FUNCTION_BLOCK logiBUS_QWA_SERVO (* Composite FB for servo word output data *)
  (* Standard: 61499-2; Description: Copyright (c) 2026 HR Agrartechnik GmbH This program and the accompanying materials are made available under the terms of the Eclipse Public License 2.0 which is available at https://www.eclipse.org/legal/epl-2.0/ SPDX-License-Identifier: EPL-2.0 *)
  (* Version 1.1, 2026-11-06, Franz Höpfinger, HR Agrartechnik GmbH, Servo on MCPWM with FREQ, PULSE_MIN, PULSE_MAX (before: LEDC, fixed 250 Hz, 800..2180 us) *)
  (* Version 1.0, 2026-02-23, Franz Höpfinger, HR Agrartechnik GmbH *)
  PACKAGE logiBUS::io::DO_SERVO;
  IMPORT logiBUS::io::DQ::logiBUS_DO::Invalid;
  IMPORT logiBUS::io::DQ::logiBUS_DO_S;
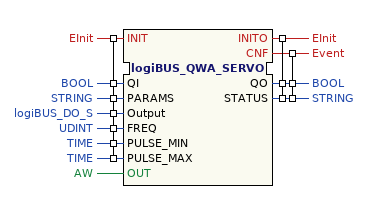
  EVENT_INPUT
    INIT : EInit WITH QI, PARAMS, Output, FREQ, PULSE_MIN, PULSE_MAX; (* Service Initialization *)
  END_EVENT
  EVENT_OUTPUT
    INITO : EInit WITH QO, STATUS; (* Initialization Confirm *)
    CNF WITH QO, STATUS; (* Confirmation of Requested Service *)
  END_EVENT
  VAR_INPUT
    QI : BOOL; (* Event Input Qualifier *)
    PARAMS : STRING; (* Service Parameters *)
    Output : logiBUS::io::DQ::logiBUS_DO_S := Invalid; (* Identify the Output Output_Q1..Q8 *)
    FREQ : UDINT := 50; (* Repetition rate of the servo pulse in Hz, read at INIT (50 Hz = one pulse every 20 ms). Servos with the same FREQ share an MCPWM timer. Standard servos 50 Hz; many car servos 250 Hz (e.g. Blue Bird BMS-L530MG: FREQ = 250, PULSE_MIN = T#1100us, PULSE_MAX = T#1900us) *)
    PULSE_MIN : TIME := T#1000us; (* Pulse width for OUT = 0, read at INIT (resolution 1 us). PULSE_MAX below PULSE_MIN turns the direction *)
    PULSE_MAX : TIME := T#2000us; (* Pulse width for OUT = 0xFAFF (100 %), read at INIT (resolution 1 us) *)
  END_VAR
  VAR_OUTPUT
    QO : BOOL; (* Event Output Qualifier *)
    STATUS : STRING; (* Service Status *)
  END_VAR
  SOCKETS
    OUT : adapter::types::unidirectional::AW; (* Servo position 0..0xFAFF (D1, 0..100 %) between PULSE_MIN and PULSE_MAX *)
  END_SOCKETS
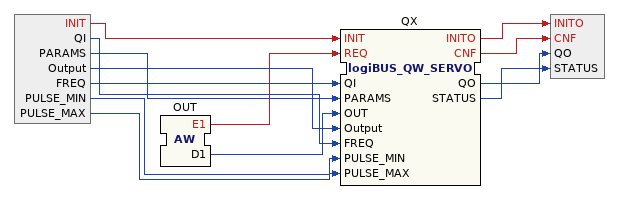
  FBS
    QX : logiBUS::io::DO_SERVO::logiBUS_QW_SERVO;
  END_FBS
  EVENT_CONNECTIONS
    INIT TO QX.INIT;
    QX.INITO TO INITO;
    OUT.E1 TO QX.REQ;
    QX.CNF TO CNF;
  END_CONNECTIONS
  DATA_CONNECTIONS
    OUT.D1 TO QX.OUT;
    QI TO QX.QI;
    PARAMS TO QX.PARAMS;
    QX.QO TO QO;
    QX.STATUS TO STATUS;
    Output TO QX.Output;
    FREQ TO QX.FREQ;
    PULSE_MIN TO QX.PULSE_MIN;
    PULSE_MAX TO QX.PULSE_MAX;
  END_CONNECTIONS
END_FUNCTION_BLOCK
